(* IEC 61131-3 sources: volt/packages/volt-lsp-iec/test-corpus/bakon-nano/Device/Plc Logic/Application/Library Manager/SysTimeCore, 4 files *)

(* ---- SYSTIME.dut ---- *)
TYPE SYSTIME : ULINT;
END_TYPE

(* ---- SYSTIMEGETMS.pou ---- *)
FUNCTION SYSTIMEGETMS : UDINT
END_FUNCTION

(* ---- SYSTIMEGETNS.pou ---- *)
FUNCTION SYSTIMEGETNS : RTS_IEC_RESULT
VAR_IN_OUT
	PUSTIME : SYSTIME;
END_VAR
END_FUNCTION

(* ---- SYSTIMEGETUS.pou ---- *)
FUNCTION SYSTIMEGETUS : RTS_IEC_RESULT
VAR_IN_OUT
	PUSTIME : SYSTIME;
END_VAR
END_FUNCTION
